FUNCTION_BLOCK FB_OnOff_Reset
(*

The function block used to activates software enable for an axis

Constructor: 		Patryk Panylo
Company:		E. Riexinger GmbH
Date:			22.09.2015
Version:			1.00

Date:			Revision:		Who:				Comment

*)
VAR_INPUT
	(* Input variables / Eingang Variablen *)
	bExecute					:BOOL;		(* Execut the function block *)
	pAxis						:POINTER TO ST_AXIS_REF_V2;
END_VAR
VAR_OUTPUT
	(* Output variables / Ausgang Variablen *)
	bDone						:BOOL;			(* Status = TRUE indicates that the axis is ready for operation. *)
	bError						:BOOL;			(* Error *)
	udnErrorNo					:UDINT;			(* Error number *)
	sErrorMsg					:STRING; 		(* Error message *)
END_VAR
VAR_IN_OUT
	(* Input Output variables / Ausgang Variablen *)

END_VAR
VAR
	(* Enummerations *)

	(* Variables *)

	(* References *)

	(* Interfaces *)

	(* Instances *)
	rtExecute						:R_TRIG;
END_VAR


rtExecute(CLK := bExecute
           		    AND pAxis^.stAxisStates.bError );       (* Error *)

IF rtExecute.Q
THEN
	pAxis^.stAxisCtrl.bFaultReset := TRUE;
END_IF;

IF NOT pAxis^.stAxisStates.bError       (* Error *)
THEN
	pAxis^.stAxisCtrl.bFaultReset := FALSE;
END_IF;

bDone := bExecute
		AND NOT  pAxis^.stAxisStates.bError;        (* Error *)

END_FUNCTION_BLOCK

(* stored: Version 1.1.0.1, ProductVersion 3.1.4024.15
   POU FB_OnOff_Reset: Id {6343e8af-f4d0-429a-a17f-7dd019c10e5e}, SpecialFunc None *)
